// TwinCAT 3 PLC project HelloWorld
// ProgramVersion: 3.1.4026.28
// libraries:
//   Tc2_Standard, * (Beckhoff Automation GmbH)
//   Tc2_System, * (Beckhoff Automation GmbH)
//   Tc3_Module, * (Beckhoff Automation GmbH)
// project tree:
//   GVLs/ IO.TcGVL
//   / PlcTask.TcTTO
//   POUs/ ExampleProgram.TcPOU, ExampleProgram2.TcPOU
// real-time tasks:
//   TASK PlcTask: cycle T#10ms, priority 20, ADS port 350
// I/O:
//   DEVICE Device 1 (EtherCAT), AmsNetId 10.169.247.170.2.1
//     Term 1 (EK1200) [EK1200-7000 EtherCAT Power supply (1,5A E-Bus)]
//       Term 2 (EL1008) [EL1008 8Ch. Dig. Input 24V, 3ms]
//       Term 3 (EL1008) [EL1008 8Ch. Dig. Input 24V, 3ms]
//       Term 4 (EL1008) [EL1008 8Ch. Dig. Input 24V, 3ms]
//       Term 5 (EL2008) [EL2008 8Ch. Dig. Output 24V, 0.5A]
//       Term 6 (EL9110) [EL9110 Power Supplier with LED (24V, Diagnostics)]
//       Term 7 (EL2008) [EL2008 8Ch. Dig. Output 24V, 0.5A]
//       Term 8 (EL7031) [EL7031 1Ch. Stepper motor output stage (24V, 1.5A)]
//       Term 9 (EL7031) [EL7031 1Ch. Stepper motor output stage (24V, 1.5A)]
//       Term 10 (EL9011) [EL9011 End Terminal]
//   DEVICE Device 2 (NOV-DP-RAM)
//   DEVICE Device 3 (CX7000), AmsNetId 10.169.247.170.4.1
//     Term 1 (CX7028) [CX7028-0000-0121]
//       modules: Module 1 (DIO_2x), Module 2 (Empty Module), Module 3 (DIO_2x), Module 4 (Empty Module), Module 5 (DI_2x), Module 6 (Empty Module), Module 7 (DI_2x), Module 8 (Empty Module)
// variable links:
//   HelloWorld/HelloWorld Instance <-> Device 1 (EtherCAT)/Term 1 (EK1200)/Term 2 (EL1008)
//     PlcTask Inputs/IO.bTerm2_In1_ModeSwitchMaintNO <-> Channel 1/Input
//     PlcTask Inputs/IO.bTerm2_In2_ModeSwitchAutoNO <-> Channel 2/Input
//     PlcTask Inputs/IO.bTerm2_In3_BtnFaultRstNO <-> Channel 3/Input
//     PlcTask Inputs/IO.bTerm2_In4_BtnFaultRstNC <-> Channel 4/Input
//     PlcTask Inputs/IO.bTerm2_In5_BtnStopRstNO <-> Channel 5/Input
//     PlcTask Inputs/IO.bTerm2_In6_BtnStopRstNC <-> Channel 6/Input
//     PlcTask Inputs/IO.bTerm2_In7_BtnParkNO <-> Channel 7/Input
//     PlcTask Inputs/IO.bTerm2_In8_BtnParkNC <-> Channel 8/Input
//   HelloWorld/HelloWorld Instance <-> Device 1 (EtherCAT)/Term 1 (EK1200)/Term 3 (EL1008)
//     PlcTask Inputs/IO.bTerm3_In1_SensStationBlk <-> Channel 1/Input
//     PlcTask Inputs/IO.bTerm3_In2_SensLiftBlk <-> Channel 2/Input
//     PlcTask Inputs/IO.bTerm3_In{3..8} <-> Channel {3..8}/Input  (6 links)
//   HelloWorld/HelloWorld Instance <-> Device 1 (EtherCAT)/Term 1 (EK1200)/Term 4 (EL1008)
//     PlcTask Inputs/IO.bTerm4_In{1..4} <-> Channel {1..4}/Input  (4 links)
//     PlcTask Inputs/IO.bTerm4_In5_BtnEStopNO <-> Channel 5/Input
//     PlcTask Inputs/IO.bTerm4_In6_BtnEStopNC <-> Channel 6/Input
//     PlcTask Inputs/IO.bTerm4_In7_BtnConfirmNO <-> Channel 7/Input
//     PlcTask Inputs/IO.bTerm4_In8_BtnConfirmNC <-> Channel 8/Input
//   HelloWorld/HelloWorld Instance <-> Device 1 (EtherCAT)/Term 1 (EK1200)/Term 5 (EL2008)
//     PlcTask Outputs/IO.bTerm5_Out1_ParkInd <-> Channel 1/Output
//     PlcTask Outputs/IO.bTerm5_Out2_ConfirmInd <-> Channel 2/Output
//     PlcTask Outputs/IO.bTerm5_Out3_StopResetInd <-> Channel 3/Output
//     PlcTask Outputs/IO.bTerm5_Out4_FaultInd <-> Channel 4/Output
//     PlcTask Outputs/IO.bTerm5_Out5_FaultResetInd <-> Channel 5/Output
//     PlcTask Outputs/IO.bTerm5_Out6_AutoModeInd <-> Channel 6/Output
//     PlcTask Outputs/IO.bTerm5_Out7_MaintModeInd <-> Channel 7/Output
//     PlcTask Outputs/IO.bTerm5_Out8_ReadyInd <-> Channel 8/Output
//   HelloWorld/HelloWorld Instance <-> Device 1 (EtherCAT)/Term 1 (EK1200)/Term 6 (EL9110)
//     PlcTask Inputs/IO.bTerm6_PowerOK <-> PowerOK/Input
//   HelloWorld/HelloWorld Instance <-> Device 1 (EtherCAT)/Term 1 (EK1200)/Term 7 (EL2008)
//     PlcTask Outputs/IO.bTerm7_Out{1..8} <-> Channel {1..8}/Output  (8 links)
//   HelloWorld/HelloWorld Instance <-> Device 3 (CX7000)/Term 1 (CX7028)
//     PlcTask Inputs/IO.bCX_In1 <-> Module 1 (DIO_2x)/DIO_2x Input Channel 1/Input
//     PlcTask Inputs/IO.bCX_In2 <-> Module 1 (DIO_2x)/DIO_2x Input Channel 2/Input
//     PlcTask Inputs/IO.bCX_In3 <-> Module 3 (DIO_2x)/DIO_2x Input Channel 1/Input
//     PlcTask Inputs/IO.bCX_In4 <-> Module 3 (DIO_2x)/DIO_2x Input Channel 2/Input
//     PlcTask Inputs/IO.bCX_In5 <-> Module 5 (DI_2x)/DI_2x Input Channel 1/Input
//     PlcTask Inputs/IO.bCX_In6 <-> Module 5 (DI_2x)/DI_2x Input Channel 2/Input
//     PlcTask Inputs/IO.bCX_In7 <-> Module 7 (DI_2x)/DI_2x Input Channel 1/Input
//     PlcTask Inputs/IO.bCX_In8 <-> Module 7 (DI_2x)/DI_2x Input Channel 2/Input
//     PlcTask Outputs/IO.bCX_Out1_EnableStopBusPwr <-> Module 1 (DIO_2x)/DIO_2x Output Channel 1/Output
//     PlcTask Outputs/IO.bCX_Out2 <-> Module 1 (DIO_2x)/DIO_2x Output Channel 2/Output
//     PlcTask Outputs/IO.bCX_Out3 <-> Module 3 (DIO_2x)/DIO_2x Output Channel 1/Output
//     PlcTask Outputs/IO.bCX_Out4 <-> Module 3 (DIO_2x)/DIO_2x Output Channel 2/Output

CONFIGURATION HelloWorld
    RESOURCE PLC ON TwinCAT3
        TASK PlcTask(INTERVAL := T#10ms, PRIORITY := 20);
        PROGRAM ExampleProgram WITH PlcTask : ExampleProgram;
        PROGRAM ExampleProgram2 WITH PlcTask : ExampleProgram2;
    END_RESOURCE
END_CONFIGURATION

// ---- GVLs/IO.TcGVL
{attribute 'qualified_only'}
VAR_GLOBAL
	// =============================================================
	// DEVICE 3: CX7000 INTEGRATED IO
	// =============================================================
	// Term 1: CX7028 Onboard Inputs (8) and Outputs (4)
	bCX_In1 AT %I* : BOOL;
	bCX_In2 AT %I* : BOOL;
	bCX_In3 AT %I* : BOOL;
	bCX_In4 AT %I* : BOOL;
	bCX_In5 AT %I* : BOOL;
	bCX_In6 AT %I* : BOOL;
	bCX_In7 AT %I* : BOOL;
	bCX_In8 AT %I* : BOOL;

	bCX_Out1_EnableStopBusPwr AT %Q* : BOOL;
	bCX_Out2 AT %Q* : BOOL;
	bCX_Out3 AT %Q* : BOOL;
	bCX_Out4 AT %Q* : BOOL;

	// =============================================================
	// DEVICE 1: ETHERCAT RAIL (EK1200)
	// =============================================================

	// Term 2: EL1008 (8 Ch. Digital Input)
	bTerm2_In1_ModeSwitchMaintNO AT %I* : BOOL;
	bTerm2_In2_ModeSwitchAutoNO AT %I* : BOOL;
	bTerm2_In3_BtnFaultRstNO AT %I* : BOOL;
	bTerm2_In4_BtnFaultRstNC AT %I* : BOOL;
	bTerm2_In5_BtnStopRstNO AT %I* : BOOL;
	bTerm2_In6_BtnStopRstNC AT %I* : BOOL;
	bTerm2_In7_BtnParkNO AT %I* : BOOL;
	bTerm2_In8_BtnParkNC AT %I* : BOOL;

	// Term 3: EL1008 (8 Ch. Digital Input)
	bTerm3_In1_SensStationBlk AT %I* : BOOL;
	bTerm3_In2_SensLiftBlk AT %I* : BOOL;
	bTerm3_In3 AT %I* : BOOL;
	bTerm3_In4 AT %I* : BOOL;
	bTerm3_In5 AT %I* : BOOL;
	bTerm3_In6 AT %I* : BOOL;
	bTerm3_In7 AT %I* : BOOL;
	bTerm3_In8 AT %I* : BOOL;

	// Term 4: EL1008 (8 Ch. Digital Input)
	bTerm4_In1 AT %I* : BOOL;
	bTerm4_In2 AT %I* : BOOL;
	bTerm4_In3 AT %I* : BOOL;
	bTerm4_In4 AT %I* : BOOL;
	bTerm4_In5_BtnEStopNO AT %I* : BOOL;
	bTerm4_In6_BtnEStopNC AT %I* : BOOL;
	bTerm4_In7_BtnConfirmNO AT %I* : BOOL;
	bTerm4_In8_BtnConfirmNC AT %I* : BOOL;

	// Term 5: EL2008 (8 Ch. Digital Output)
	bTerm5_Out1_ParkInd AT %Q* : BOOL;
	bTerm5_Out2_ConfirmInd AT %Q* : BOOL;
	bTerm5_Out3_StopResetInd AT %Q* : BOOL;
	bTerm5_Out4_FaultInd AT %Q* : BOOL;
	bTerm5_Out5_FaultResetInd AT %Q* : BOOL;
	bTerm5_Out6_AutoModeInd AT %Q* : BOOL;
	bTerm5_Out7_MaintModeInd AT %Q* : BOOL;
	bTerm5_Out8_ReadyInd AT %Q* : BOOL;

	// Term 6: EL9110 (Power Feed with Diagnostics)
	bTerm6_PowerOK      AT %I* : BOOL; // True if the 24V bus is healthy

	// Term 7: EL2008 (8 Ch. Digital Output)
	bTerm7_Out1 AT %Q* : BOOL;
	bTerm7_Out2 AT %Q* : BOOL;
	bTerm7_Out3 AT %Q* : BOOL;
	bTerm7_Out4 AT %Q* : BOOL;
	bTerm7_Out5 AT %Q* : BOOL;
	bTerm7_Out6 AT %Q* : BOOL;
	bTerm7_Out7 AT %Q* : BOOL;
	bTerm7_Out8 AT %Q* : BOOL;

	// Term 8: EL7031 (Stepper Motor Drive)
	nTerm8_Status  AT %I* : UINT;
	nTerm8_Pos     AT %I* : UDINT;
	nTerm8_Control AT %Q* : UINT;
	nTerm8_Velo    AT %Q* : INT;

	// Term 9: EL7031 (Stepper Motor Drive)
	nTerm9_Status  AT %I* : UINT;
	nTerm9_Pos     AT %I* : UDINT;
	nTerm9_Control AT %Q* : UINT;
	nTerm9_Velo    AT %Q* : INT;

	// Term 10: EL9011 (End Cap)
	// (No logic mapping; it's just a piece of plastic.)

END_VAR

// ---- POUs/ExampleProgram.TcPOU
PROGRAM ExampleProgram
VAR
END_VAR

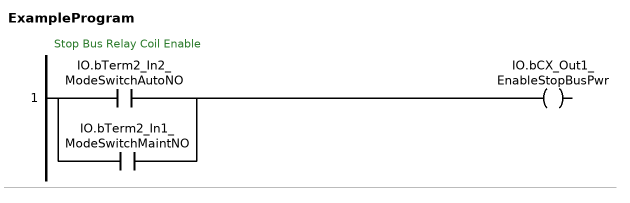
// NETWORK 1
// Stop Bus Relay Coil Enable
IO.bCX_Out1_EnableStopBusPwr := IO.bTerm2_In2_ModeSwitchAutoNO OR IO.bTerm2_In1_ModeSwitchMaintNO;

END_PROGRAM

// ---- POUs/ExampleProgram2.TcPOU
PROGRAM ExampleProgram2
VAR
	fbTimerOff  : TON;
    fbTimerOn   : TON;
    tOffTime    : TIME := T#1000MS; // Mappable off-time
    tOnTime     : TIME := T#1000MS; // Mappable on-time
    bBlinkerOn  : BOOL;
	bBlinkerOff : BOOL;
END_VAR

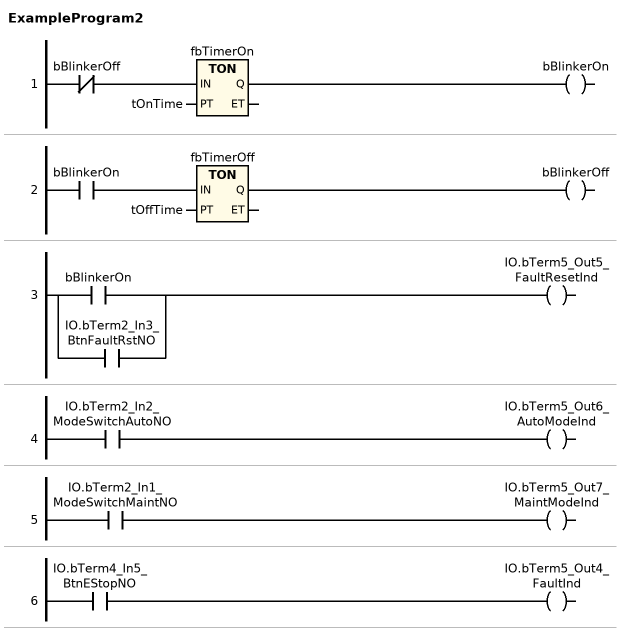
// NETWORK 1
fbTimerOn(IN := NOT bBlinkerOff, PT := tOnTime); // TON
bBlinkerOn := fbTimerOn.Q;

// NETWORK 2
fbTimerOff(IN := bBlinkerOn, PT := tOffTime); // TON
bBlinkerOff := fbTimerOff.Q;

// NETWORK 3
IO.bTerm5_Out5_FaultResetInd := bBlinkerOn OR IO.bTerm2_In3_BtnFaultRstNO;

// NETWORK 4
IO.bTerm5_Out6_AutoModeInd := IO.bTerm2_In2_ModeSwitchAutoNO;

// NETWORK 5
IO.bTerm5_Out7_MaintModeInd := IO.bTerm2_In1_ModeSwitchMaintNO;

// NETWORK 6
IO.bTerm5_Out4_FaultInd := IO.bTerm4_In5_BtnEStopNO;

END_PROGRAM
